// TIA Portal V20 export
// export: Created 2026-10-12T16:46:22.7186029Z, ExportSetting WithDefaults, DisplayName Totally Integrated Automation Portal, DisplayVersion V20 Update 6, DisplayName TIA Portal Openness, DisplayVersion V20 Update 6, DisplayName TIA Portal Version Control Interface, DisplayVersion V20 Update 6, DisplayName SINAMICS Startdrive Advanced, DisplayVersion V20 SP1 Update 2, DisplayName SINAMICS Startdrive G110M, G120, G120C, G120D, G120P, G115D, DisplayVersion V20 SP1 Update 2, DisplayName SINAMICS Startdrive G130, G150, S120, S150, SINAMICS MV, G220, S200, S210, DisplayVersion V20 SP1 Update 2, DisplayName STEP 7 Professional, DisplayVersion V20 Update 6, DisplayName STEP 7 Safety, DisplayVersion V20 Update 2, DisplayName WinCC Basic/Comfort/Advanced, DisplayVersion V20 Update 6, DisplayName WinCC Professional, DisplayVersion V20 Update 6, DisplayName WinCC Unified, DisplayVersion V20 Update 6
TYPE "UDT_FlexKraft_Out"
// ==============================================================================
//   FlexKraft via Anybus Communicator (PROFINET)  -  SCL-Quelldatei
// ------------------------------------------------------------------------------
//   Erzeugt 3 UDTs, 1 globalen DB und 1 FB:
//       UDT_FlexKraft_Out      (32 Byte, SPS  -> FK Holding-Register 0..15)
//       UDT_FlexKraft_In       (32 Byte, FK Input-Register 0..15  -> SPS)
//       UDT_FlexKraft_Device   (Wrapper Out + In, 64 Byte)
//       DB_FlexKraft_Data      (3 x Device  -> FK_1, FK_2, FK_3)
//       FB_FlexKraft           (Komfort-Bitzerlegung des Control-/Statusworts)
// 
//   Voraussetzungen:
//     - Anybus Communicator (PROFINET-Firmware) als IO-Device in TIA eingebunden
//     - I/O-Map gemÃ¤ÃŸ Gateway-Export:
//           FK_1  Modbus 2  Bytes  0..31
//           FK_2  Modbus 3  Bytes 32..63
//           FK_3  Modbus 4  Bytes 64..95
//     - FK im Output Mode "Series/Parallel"; bei Dual-Mode UDT-Layout anpassen
//     - Am Gleichrichter: PROTOCOL=MODBUS RTU, POWERONMODE=Remote, eindeutige Adr.
// 
//   Wichtig zum Datenaustausch:
//     - DB ist mit "Optimierter Bausteinzugriff = FALSE" deklariert, damit das
//       Byte-Layout vorhersagbar ist und ein direkter Word-Copy aus/in die
//       Peripherie mÃ¶glich ist. Beispiel-OB1-Snippet ganz unten.
//     - Als sichere Alternative bei optimierten Bausteinen:
//       DPRD_DAT / DPWR_DAT mit der HW-Kennung des Submoduls.
// ==============================================================================
// ==============================================================================
//  UDT 1: Output (SPS -> Gateway -> FK Holding Register 0..15)
// ==============================================================================
// stored: IsFailsafeCompliant false
   STRUCT
      PageNo : Word;   // Reg 0 reserviert, immer 16#0000
      ControlRegister : Word;   // Reg 1 Bitfeld, siehe FB / Bittabelle
      SetVoltage : Int;   // Reg 2 Sollspannung *0,01 V (signed)
      SetCurrent : Int;   // Reg 3 Sollstrom *1 A bzw. *0,1 A (HiRes)
      ProcessTimerLimit_HW : Word;   // Reg 4 *65535 s
      ProcessTimerLimit_LW : Word;   // Reg 5 *1 s
      AhLimit_HW : Word;   // Reg 6 *65536 Ah
      AhLimit_LW : Word;   // Reg 7 *1 Ah
      Startramp : Word;   // Reg 8 Anlauframpe *0,1 s
      Reserved : Array[9..15] of Word;   // Reg 9..15 ungenutzt
   END_STRUCT;
END_TYPE
